SUBAPPLICATION Uebung_269_AX (* Dialog: Toast (Hinweis ohne Tasten, verschwindet nach 3 s), Pool Dialog *)
  (* Standard: 61499-2; Description: Copyright (c) 2026 Meisterschulen am Ostbahnhof This program and the accompanying materials are made available under the terms of the Eclipse Public License 2.0 which is available at https://www.eclipse.org/legal/epl-2.0/ SPDX-License-Identifier: EPL-2.0 *)
  (* Version 1.0, 2026-11-17, Franz Höpfinger, Meisterschulen am Ostbahnhof, initial API and implementation and/or initial documentation *)
  PACKAGE Uebungen;
  IMPORT Uebungen::const::UT::Dialog::DefaultPool::OutputString_Text_Toast;
  IMPORT Uebungen::const::UT::Dialog::DefaultPool::SoftKey_F1;
  IMPORT isobus::UT::dialog::DialogConst::DLG_ICON_INFO;
  IMPORT isobus::UT::io::Softkey::SoftKeyActivationCode::SK_RELEASED;
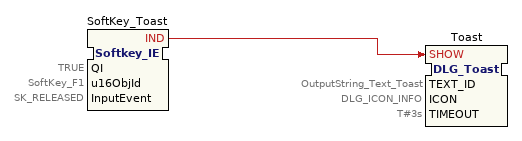
  FBS
    SoftKey_Toast : isobus::UT::io::Softkey::Softkey_IE(QI := TRUE, u16ObjId := SoftKey_F1, InputEvent := SK_RELEASED);
    Toast : isobus::UT::dialog::DLG_Toast(TEXT_ID := OutputString_Text_Toast, ICON := DLG_ICON_INFO, TIMEOUT := T#3s);
  END_FBS
  EVENT_CONNECTIONS
    SoftKey_Toast.IND TO Toast.SHOW;
  END_CONNECTIONS
END_SUBAPPLICATION
